{attribute 'qualified_only'}
VAR_GLOBAL
    {attribute 'OPC.UA.DA' := '1'}
    nIn  : DINT;   // escrito pelo cliente (Python)
    {attribute 'OPC.UA.DA' := '1'}
    nOut : DINT;   // eco: PRG_Echo copia nIn aqui a cada ciclo
END_VAR

(* stored: Version 1.1.0.1, ProductVersion 3.1.4026.0
   GVL GVL_Bench: Id {4d1c0a52-7b0e-4a41-9b6e-0c1d5e7a2f01} *)
